(* PLC project g_hvac_fan_delay_bomb, Anonymous Benchmark Suite 1.0 *)
(* stored: creationDateTime 2026-07-09T00:00:00 *)

PROGRAM g_hvac_fan_delay_bomb
  VAR_INPUT
    heat_call : BOOL;
    cool_call : BOOL;
    enable : BOOL;
    maint : BOOL;
  END_VAR
  VAR_OUTPUT
    heat : BOOL;
    cool : BOOL;
    fan : BOOL;
  END_VAR

(* LD diagram, written out as Structured Text *)
heat := (NOT cool_call OR cool_call AND maint) AND heat_call AND enable;
cool := cool_call AND enable;
fan := enable;
END_PROGRAM

CONFIGURATION Config0
  RESOURCE Res0 ON PLC
    TASK tcyclic(INTERVAL := T#10ms, PRIORITY := 0);
    PROGRAM inst0 WITH tcyclic : g_hvac_fan_delay_bomb;
  END_RESOURCE
END_CONFIGURATION
